// Größte zulässige Z1-Position (Futter <-> Führung) bei gegebener Z2-Position.
FUNCTION F_Z1Max : LREAL
VAR_INPUT
    fZ2 : LREAL;
END_VAR

F_Z1Max := GVL_Config.fZ1CollisionBase_mm + fZ2;

END_FUNCTION

(* stored: Version 1.1.0.1
   POU F_Z1Max: Id {53b0a940-1f15-594a-87fe-156330e62e2c}, SpecialFunc None *)
